{attribute 'qualified_only'}
{attribute 'strict'}
{attribute 'to_string'}
TYPE E_ModuleState :
(
	Unknown 	:= 0,
	Starting 	:= 1,
	Started		:= 2,
	Stopping	:= 4,
	Stopped		:= 8
) INT;
END_TYPE

(* stored: Version 1.1.0.1, ProductVersion 3.1.4024.12
   DUT E_ModuleState: Id {0f3ea25b-dee5-4489-bf2a-4bd07d76c5d3} *)
